FUNCTION_BLOCK Model (* Composite Function Block Type *)
  (* Standard: 61499-2 *)
  (* Version 0.0, 6/20/2016, Andrei, nxtControl GmbH, template *)
  PACKAGE Main;
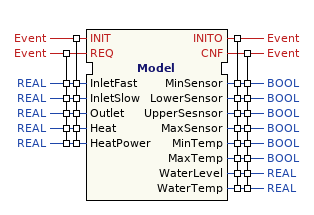
  EVENT_INPUT
    INIT WITH InletFast, InletSlow, Outlet, Heat, HeatPower; (* Initialization Request *)
    REQ WITH InletFast, InletSlow, Outlet, Heat, HeatPower; (* Normal Execution Request *)
  END_EVENT
  EVENT_OUTPUT
    INITO WITH MinSensor, LowerSensor, UpperSesnsor, MaxSensor, MinTemp, MaxTemp, WaterLevel, WaterTemp; (* Initialization Confirm *)
    CNF WITH MinSensor, LowerSensor, UpperSesnsor, MaxSensor, MinTemp, MaxTemp, WaterLevel, WaterTemp; (* Execution Confirmation *)
  END_EVENT
  VAR_INPUT
    InletFast : REAL; (* Input event qualifier *)
    InletSlow : REAL;
    Outlet : REAL;
    Heat : REAL;
    HeatPower : REAL;
  END_VAR
  VAR_OUTPUT
    MinSensor : BOOL; (* Output event qualifier *)
    LowerSensor : BOOL;
    UpperSesnsor : BOOL;
    MaxSensor : BOOL;
    MinTemp : BOOL;
    MaxTemp : BOOL;
    WaterLevel : REAL;
    WaterTemp : REAL;
  END_VAR
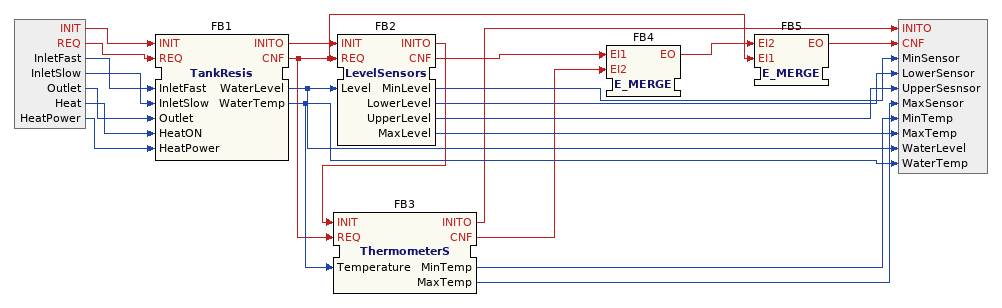
  FBS
    FB1 : TankResis;
    FB4 : E_MERGE;
    FB3 : ThermometerS;
    FB2 : LevelSensors;
    FB5 : E_MERGE;
  END_FBS
  EVENT_CONNECTIONS
    FB3.INITO TO INITO;
    INIT TO FB1.INIT;
    REQ TO FB1.REQ;
    FB1.INITO TO FB2.INIT;
    FB1.CNF TO FB2.REQ;
    FB2.INITO TO FB3.INIT;
    FB1.CNF TO FB3.REQ;
    FB2.CNF TO FB4.EI1;
    FB5.EO TO CNF;
    FB3.CNF TO FB4.EI2;
    FB4.EO TO FB5.EI2;
    FB1.CNF TO FB5.EI1;
  END_CONNECTIONS
  DATA_CONNECTIONS
    FB2.MinLevel TO MinSensor;
    FB2.LowerLevel TO LowerSensor;
    FB2.UpperLevel TO UpperSesnsor;
    FB2.MaxLevel TO MaxSensor;
    FB3.MinTemp TO MinTemp;
    FB3.MaxTemp TO MaxTemp;
    FB1.WaterLevel TO FB2.Level;
    InletFast TO FB1.InletFast;
    InletSlow TO FB1.InletSlow;
    Outlet TO FB1.Outlet;
    Heat TO FB1.HeatON;
    FB1.WaterTemp TO FB3.Temperature;
    FB1.WaterTemp TO WaterTemp;
    FB1.WaterLevel TO WaterLevel;
    HeatPower TO FB1.HeatPower;
  END_CONNECTIONS
END_FUNCTION_BLOCK
